(* IEC 61131-3 sources: plc-ci-toolkit/tools/tests/fixtures/sourcemap/src/GVLs, 1 file *)

(* ---- GVL_Const.gvl.st ---- *)
// Пример для проверки карты строк после понижения iec-checker (tools/tests): метка @N в комментарии —
// номер строки в этом файле; сравнения с 1.5 в условиях IF дают PLCOPEN-CP8
VAR_GLOBAL CONSTANT
    SLOTS_MAX : INT := 4;    // @4
    NAME_SIZE : INT := 16;   // @5
END_VAR
